Fanuc KAREL source: KO00048.KL

PROGRAM KO00048
%NOLOCKGROUP
%ENVIRONMENT MIR
VAR
  P1: POSITION
  P2: JOINTPOS
  F: BOOLEAN
  OUT: JOINTPOS
BEGIN
  F = TRUE
  OUT = MIRROR(P1, P2, F)
END KO00048
